(* IEC 61131-3 sources: Versio-VersionControlSystem/fixtures/projects/TC3_PlcSample_reStrText/TC3_PlcSample_reStrText/LibraryDocumentationSample Project/LibPOUs/B_DocuElements/Hyperlinks, 7 files *)

(* ---- FB_Libdoc_AnonymousHyperlinks.st ---- *)
(*
See the `Beckhoff Online Information System`__ or the `Beckhoff home page`__.

.. __: http://infosys.beckhoff.de/

.. __: http://beckhoff.de/
*)

FUNCTION_BLOCK FB_Libdoc_AnonymousHyperlinks
VAR_INPUT
    nVarA : INT;
    nVarB : INT;
END_VAR
VAR_OUTPUT
    nSum : INT;
END_VAR
VAR
END_VAR

(* ---- FB_Libdoc_Citation.st ---- *)
(*
Citation references, like [CIT2002]_. Note that citations may get rearranged, e.g., to the bottom of the "page".

| Some sample text to get some text in between.
| Some sample text to get some text in between.
| Some sample text to get some text in between.
| Some sample text to get some text in between.
| Some sample text to get some text in between.
| Some sample text to get some text in between.

.. [CIT2002] This is the citation.  It's just like a footnote,
   except the label is textual.

Given a citation like [this]_, one can also refer to it like this_.

| Some sample text to get some text in between.
| Some sample text to get some text in between.
| Some sample text to get some text in between.
| Some sample text to get some text in between.
| Some sample text to get some text in between.
| Some sample text to get some text in between.

.. [this] here.

| Some sample text to get some text in between.
| Some sample text to get some text in between.
| Some sample text to get some text in between.
| Some sample text to get some text in between.
| Some sample text to get some text in between.
| Some sample text to get some text in between.

*)

FUNCTION_BLOCK FB_Libdoc_Citation
VAR_INPUT
    nVarA : INT;
    nVarB : INT;
END_VAR
VAR_OUTPUT
    nSum : INT;
END_VAR
VAR
END_VAR

(* ---- FB_Libdoc_ExternalHyperlinks.st ---- *)
(*
See the Beckhoff homepage_ for more information.

Please contact the `Beckhoff Support`_ for technical assistance.

.. _homepage: http://www.beckhoff.de
.. _Beckhoff Support: support@beckhoff.com

For more information see the `PLC Lib Tc2_System`_ and `PLC Lib Tc2_Standard`_.

.. _PLC Lib Tc2_System: https://download.beckhoff.com/download/document/automation/twincat3/TwinCAT_3_PLC_Lib_Tc2_System_EN.pdf
.. _PLC Lib Tc2_Standard: https://download.beckhoff.com/download/document/automation/twincat3/TwinCAT_3_PLC_Lib__Tc2_Standard_EN.pdf

External hyperlinks, like `Beckhoff <http://www.beckhoff.de/>`_.

**Standalone hyperlinks**

See http://www.beckhoff.de for info.

Contact support@beckhoff.com

**Embedded URIs and aliases**

See the `Beckhoff homepage <http://www.beckhoff.de>`_ for info.

This `link <Beckhoff homepage_>`_ is an alias to the link above.

See the `Beckhoff homepage`_ for info.

This link_ is an alias to the link above.

.. _Beckhoff homepage: http://www.beckhoff.de
.. _link: `Beckhoff homepage`_

*)

FUNCTION_BLOCK FB_Libdoc_ExternalHyperlinks
VAR_INPUT
    nVarA : INT;
    nVarB : INT;
END_VAR
VAR_OUTPUT
    nSum : INT;
END_VAR
VAR
END_VAR

(* ---- FB_Libdoc_IndirectHyperlinks.st ---- *)
(*

**Indirect references to an internal reference target**

This hyperlink points to target one_ and indirect to target three.

.. _one: two_
.. _two: three_
.. _three:

The hyperlink targets above point to this paragraph.

**Indirect references to an external reference target**

The `Beckhoff Information System`_ is a reference source for Beckhoff_ products

.. _Beckhoff: `Beckhoff Information System`_

.. _Beckhoff Information System: https://infosys.beckhoff.de/
*)

FUNCTION_BLOCK FB_Libdoc_IndirectHyperlinks
VAR_INPUT
    nVarA : INT;
    nVarB : INT;
END_VAR
VAR_OUTPUT
    nSum : INT;
END_VAR
VAR
END_VAR

(* ---- FB_Libdoc_InlineHyperlinks.st ---- *)
(*
| This function block is based on a _`statemachine` concept which is described in the following.
| The statemachine is based on several states.
| The proceeding always begins in the first state.
| If the last state is left, the execution restarts in the first state.
| There are so many more information necessary to describe the statemachine concept in detail.
| But as this is just a sample text to show the inline hyperlinks, we want to leave out the details.
| A rough description should be enough for the sample demonstration.
|
| Some sample text to get some text in between.
| Some sample text to get some text in between.
| Some sample text to get some text in between.
| Some sample text to get some text in between.
| Some sample text to get some text in between.
| Some sample text to get some text in between.
|
| Furthermore, the function block is based on another concept. This is called XY.
| It is always necessary to respect the demands of this concept.
| Especially, as it is deeply interwoven with the statemachine concept.
| Therefore, you definitely need to understand the statemachine concept first.
| Afterwards, you might understand the XY concept.
| For more information about this, see the description of the `statemachine`_.
| By clicking on this link, the Library Manager will jump to the beginning of the first paragraph where the statemachine concept is described..

*)

FUNCTION_BLOCK FB_Libdoc_InlineHyperlinks
VAR_INPUT
    nVarA : INT;
    nVarB : INT;
END_VAR
VAR_OUTPUT
    nSum : INT;
END_VAR
VAR
END_VAR

(* ---- FB_Libdoc_InternalHyperlinks.st ---- *)
(*

**Simple internal hyperlink target**

Clicking on this internal hyperlink will take us to the target_
below.

.. _target:

**Nesting of internal hyperlink targets**

Clicking on this internal hyperlink will take us to the `third item`_ of the bullet list.

* First list item
* Second list item

  .. _third item:

* Third list item, with hyperlink target.

**Concatentation of internal hyperlink targets**

Clicking on this internal hyperlink will take us to target1_
and clicking on this internal hyperlink will take us to target2_.
Both targets point the the same paragraph.

.. _target1:
.. _target2:

The targets "target1" and "target2" are synonyms; they both
point to this paragraph.
*)

FUNCTION_BLOCK FB_Libdoc_InternalHyperlinks
VAR_INPUT
    nVarA : INT;
    nVarB : INT;
END_VAR
VAR_OUTPUT
    nSum : INT;
END_VAR
VAR
END_VAR

(* ---- FB_Libdoc_LinkToAnotherObject.st ---- *)
(*
| It is also possible to create a reference to the documentation of another object which is also part of this library.
| For example, by clicking on this link :ref:`FB_Libdoc_InlineHyperlinks`, the documentation of this FB will be shown.
| Or you can also create a link to :ref:`FB_Libdoc_CodeBlock` which is part of another folder.

*)

FUNCTION_BLOCK FB_Libdoc_LinkToAnotherObject
VAR_INPUT
    nVarA : INT;
    nVarB : INT;
END_VAR
VAR_OUTPUT
    nSum : INT;
END_VAR
VAR
END_VAR
